Yaskawa INFORM job: CIRCLE.JBI

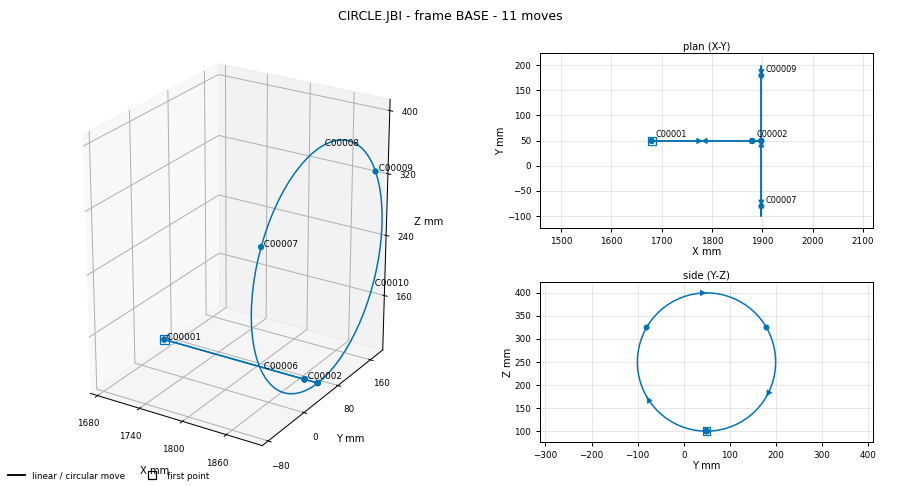
[picture p0: tool path of CIRCLE.JBI in frame BASE, 11 of 15 moves have a stored position in this frame; points joined in program order, loops and branches not executed]
/JOB
//NAME CIRCLE
//POS
///NPOS 15,0,0,0,0,0
///TOOL 9
///POSTYPE PULSE
///PULSE
C00000=2,16,-49,-2,65,91
///TOOL 9
///POSTYPE BASE
///RECTAN
///RCONF 1,0,0,0,0,0,0,0
C00001=1680.000,49.386,100.000,90.00,-0.00,90.00
C00002=1880.000,49.386,100.000,90.00,-0.00,90.00
C00003=1880.000,49.386,100.000,90.00,-0.00,90.00
C00004=1898.000,49.386,100.000,90.00,-0.00,90.00
C00005=1898.000,49.386,100.000,90.00,-0.00,90.00
C00006=1898.000,-80.510,174.986,90.00,-0.00,90.00
C00007=1898.000,-80.534,324.973,90.00,-0.00,90.00
C00008=1898.000,49.386,400.000,90.00,-0.00,90.00
C00009=1898.000,179.306,324.973,90.00,0.00,90.00
C00010=1898.000,179.282,174.986,90.00,0.00,90.00
C00011=1898.000,49.386,100.000,90.00,-0.00,90.00
C00012=1880.000,49.386,100.000,90.00,-0.00,90.00
C00013=1880.000,49.386,100.000,90.00,-0.00,90.00
C00014=1680.000,49.386,100.000,90.00,-0.00,90.00
//INST
///DATE 2026/10/26 01:19
///COMM Generated using RoboDK
///ATTR SC,RW,RJ
///GROUP1 RB1
NOP
'Using Tool2 (targets wrt base
'):
'1900.0,49.4,250.0,90.0,0.0,-9
'0.0
'Setting Tool 9 (USER - ENGRAV
'E - 30 DEG POINT END):
SETE P00095 (1) 0
SETE P00095 (2) 0
SETE P00095 (3) 85000
SETE P00095 (4) 0
SETE P00095 (5) 0
SETE P00095 (6) 0
SETTOOL TL#(9) P00095
'hide BALL END - 10MM
'show USER - ENGRAVE - 30 DEG
'POINT END
MSG "/ ALPHACAM DRAWING FILE -"
MSG " ROBOTAPT"
MSG "/ NC CODE FILE - ROBOTAPT"
MSG ".apt"
MSG "/ POST-PROCESSED FOR APT-"
MSG "CL DATA"
MSG "/ CREATED - 26 NOV 18"
MSG "/ PROGRAMMED BY ALPHACAM"
MSG "/ USER - ENGRAVE - 30 DEG"
MSG " POINT END"
MOVJ C00000 VJ=50.00
MOVL C00001 V=1000.0
MOVL C00002 V=1000.0
CALL JOB:SPINDLE
MOVL C00003 V=1000.0
MOVL C00004 V=166.7
MOVC C00005 V=166.0
MOVC C00006 V=166.0
MOVC C00007 V=166.0
MOVC C00008 V=166.7
MOVC C00009 V=166.7
MOVC C00010 V=166.7
MOVC C00011 V=166.7
MOVL C00012 V=1000.0
CALL JOB:SPINDLE
MOVL C00013 V=1000.0
MOVL C00014 V=1000.0
END
